// Mitsubishi GX Works2 project: Task2_Ex_1   PLC: FX3G

PROGRAM MAIN
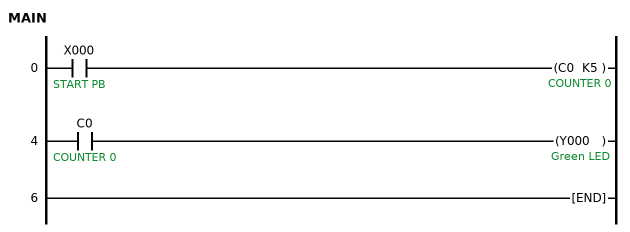
0     LD      X000  ; START PB
      OUT     C0 K5  ; COUNTER 0
4     LD      C0  ; COUNTER 0
      OUT     Y000  ; Green LED
6     END
END_PROGRAM
